Fanuc KAREL source: KT00535.KL

PROGRAM KT00535
%NOLOCKGROUP
VAR
  P1: JOINTPOS
  P2: POSITION
  OUT: XYZWPR
BEGIN
  OUT = P1 : P2
END KT00535
